ABB RobotStudio station: NeuralGrasp.rsstn

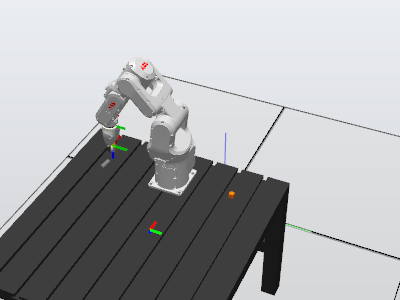
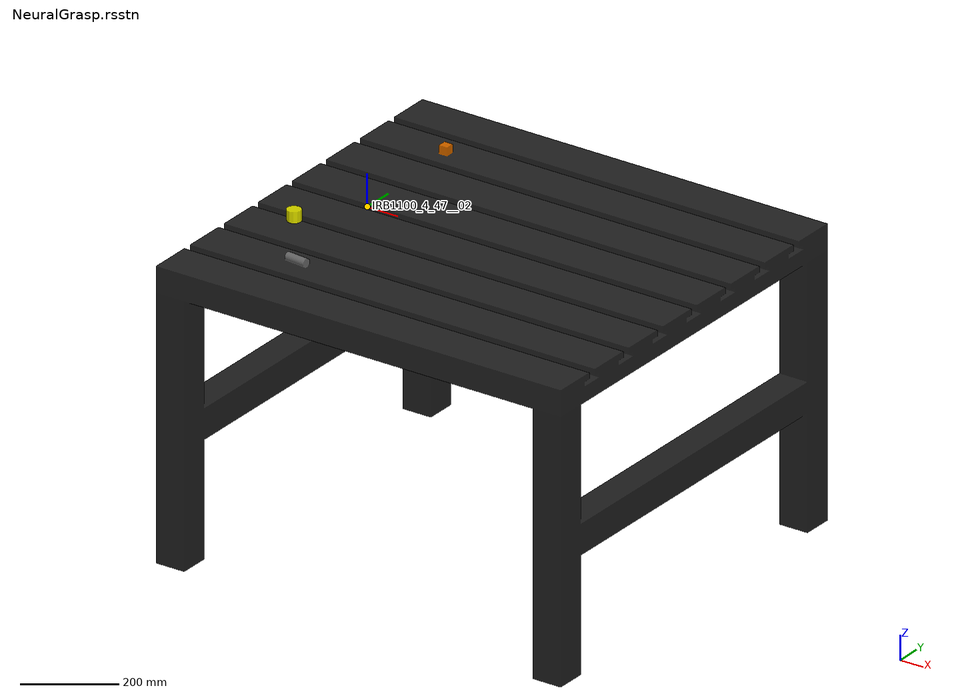
[picture v1: parts stored in the station drawn from their meshes, with robot base, taught points and paths (robot models come from the ABB library and are not in the file)]
Station NeuralGrasp (saved by RobotStudio 26.3.11844.1)
Controller ControllerC30, task T_ROB1: task frame (RAPID world) sits at (607.14, 0, 668.57) mm in the station
Controller ControllerC30
  mechanical unit ROB_1: IRB1100_4_47__02, 6 joints, base frame (0, 0, 0) mm
Layout (positions relative to the parent item):
  - IRB1100_4_47__02 [mechanism, from %ABB.RobotStudio.Models.IRB1100%\IRB1100_4_47__02.rslib] at (607.14, 0, 668.57) mm; joint values [-1.518, 0.6948, 0.3424, 0, 0.5337, -1.518] (rad or m)
  - tGrasp [mechanism, from %ABB.RobotStudio.Models.SmartGripper%\ABB_Smart_Gripper_Servo_Fingers.rslib] at (621.91, -279.44, 894.26) mm, rotated rx -180 ry 0 rz 180 deg; joint values [0.025] (rad or m)
  - Table AW Training [part] at (755.1, 0, 141.41) mm, size 1000 x 940 x 668 mm
  - box [part] at (-324.96, 215.82, 8.26) mm, size 20 x 20 x 20 mm
  - cylinder [part] at (943.29, 590.05, 15.04) mm, rotated rx 0 ry 0 rz -96.37 deg, size 20 x 50 x 19.9 mm
  - Gripper [smart component]
      signals: DI Open, DI Close
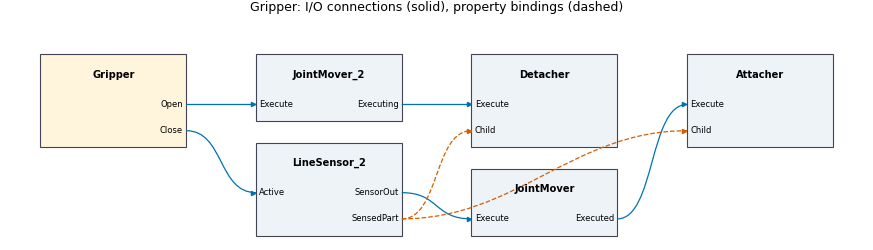
      connections:
        Gripper.Open -> JointMover_2.Execute
        JointMover_2.Executing -> Detacher.Execute
        JointMover.Executed -> Attacher.Execute
        Gripper.Close -> LineSensor_2.Active
        LineSensor_2.SensorOut -> JointMover.Execute
        LineSensor_2.SensedPart => Attacher.Child
        LineSensor_2.SensedPart => Detacher.Child
    - Attacher [smart component, from Components\Attacher.rslib]
        properties: Parent=tGrasp; Flange=0; Child=cylinder; Mount=false; Offset=[0 0 0]; Orientation=[0 0 0]
    - Detacher [smart component, from Components\Detacher.rslib]
        properties: Child=cylinder; KeepPosition=true
    - JointMover [smart component, from Components\JointMover.rslib]
        properties: Mechanism=tGrasp; Relative=false; Duration=1; J1=0.012
    - JointMover_2 [smart component, from Components\JointMover.rslib]
        properties: Mechanism=tGrasp; Relative=false; Duration=1; J1=0.025
    - LineSensor_2 [smart component, from Components\LineSensor.rslib] at (621.91, -279.44, 780.06) mm, rotated rx -180 ry 0 rz 180 deg
        properties: Start=[0 0 0]; End=[0 0 0.025]; Length=0.025; Radius=0.016; Tag=(none); SenseMultiple=false; SensedPart=cylinder; SensedPoint=[0.8859737548828125 -0.02365008544921875 0.6855578002929688]
      - _sensorPart_ [part], size 32 x 32 x 25 mm
Attachment: tGrasp is attached to IRB1100_4_47__02 / Link6
Attachment: LineSensor_2 is attached to tGrasp / HandBase
Station logic (signal -> signal, property => property):
  ControllerC30.do_Gripper -> SmartComponent_1.di_Grasp
  ControllerC30.GripperOpen -> Gripper.Open
  ControllerC30.GripperClose -> Gripper.Close
Targets, tools, work objects and paths stored in the station, written as RAPID:
! task T_ROB1
MODULE CalibData
  PERS tooldata Servo:=[TRUE,[[0,0,114.2],[1,0,0,0]],[0.215,[8.7,12.3,49.2],[1,0,0,0],0.00021,0.00024,0.00009]];
ENDMODULE

! task T_ROB1
MODULE Module1
  CONST robtarget Target_box:=[[323.849178583,62.404,20.842552413],[0,0,1,0],[0,0,0,0],[9E+09,9E+09,9E+09,9E+09,9E+09,9E+09]];
  PROC Path_10()
  ENDPROC
ENDMODULE

